(*
SPDX-FileCopyrightText: © 2026 Oleksandr Tiutyk <trofimich@gmail.com>
SPDX-License-Identifier: MIT
License: https://opensource.org/license/mit
*)

(*!
<summary>Represents a named event occurrence without additional payload.</summary>
<description>
Copies its initialization name into instance storage and exposes it through the read-only INamed contract. The
caller must supply a nonempty name. Global uniqueness is not required; each recipient defines how it
recognizes events. Equal names alone do not establish event instance identity. The Event lifetime contract
applies: one instance per occurrence, synchronous borrowed delivery, no retention by recipients and no reset
for reuse as another occurrence. Heap allocation is not required.
</description>
*)

{attribute 'no_explicit_call' := 'do not call this function block directly'}
FUNCTION_BLOCK SimpleEvent EXTENDS Event IMPLEMENTS INamed
VAR_STAT
	//! <summary>Class name shared by all instances of this function block.</summary>
	{attribute 'hide'} 
	_ClassName : STRING := __POUNAME();
END_VAR
VAR
	{attribute 'hide'} 
	_Name : WSTRING;
END_VAR

{attribute 'monitoring' := 'call'}
PROPERTY ClassName : REFERENCE TO STRING
GET
ClassName REF= _ClassName;
END_GET
END_PROPERTY

(*!
<summary>Initializes the event's name; Event initialization associates the optional source.</summary>
<description>
Copies the name into instance storage. The source is borrowed without ownership transfer; the caller must keep
a non-null source alive for the entire event lifetime. The caller must supply a nonempty name; this
precondition is not checked at runtime. Pass both additional initialization arguments explicitly; zero is
allowed for sourceObject.
</description>
*)

//!<param name="sourceObject">Source of the event, or 0 for an event without a specific source.</param>
//!<param name="name">Nonempty name copied into this event instance; global uniqueness is not required.</param>
METHOD FB_init : BOOL
VAR_INPUT
	bInitRetains : BOOL; // TRUE: the retain variables are initialized (reset warm / reset cold)
	bInCopyCode : BOOL;  // TRUE: the instance will be copied to the copy code afterward (online change)
	sourceObject : IObject;
	name : WSTRING;
END_VAR
_Name := name;
END_METHOD

(*!
<summary>Returns a borrowed, read-only view of the event's nonempty name.</summary>
<description>
Requires initialization with a nonempty name. The reference remains usable only while this instance is alive;
callers must not write through it. Recognition rules belong to the recipient, and names need not be globally
unique.
</description>
*)

{attribute 'monitoring' := 'call'}
PROPERTY FINAL Name : REFERENCE TO WSTRING
GET
Name REF= _Name;
END_GET
END_PROPERTY

(*!
<summary>Provides the library namespace used in diagnostics.</summary>
<description>
Borrowed read-only reference to the compiler-initialized library namespace; no ownership transfer.
</description>
*)
{attribute 'monitoring' := 'call'}
PROPERTY NamespaceName : REFERENCE TO STRING
GET
NamespaceName REF= CurrentNamespace.Name;
END_GET
END_PROPERTY

(*!
<summary>Reports the byte size of this concrete instance.</summary>
<description>
Uses XSIZEOF on the instance. Does not include separately allocated payloads or prove that an arbitrary
address is valid.
</description>
*)
{attribute 'monitoring' := 'call'}
PROPERTY SelfSize : ULINT
GET
SelfSize := XSIZEOF(THIS^);
END_GET
END_PROPERTY

END_FUNCTION_BLOCK

(* stored: Version 1.1.0.1
   POU SimpleEvent: Id {6068111a-5f7a-4513-bc9f-2ae69d62cec9}, SpecialFunc None
   Property ClassName: Id {74c80bc7-04ea-415b-b755-fddcf5a7aecd}
   Get Get: Id {0b51e612-0055-4cf8-b992-12a817738a31}
   Method FB_init: Id {95fe79f8-57ab-4f8f-8458-df22c083e6ed}
   Property Name: Id {4cc1da98-6df4-40c6-a0ac-2b058bef2a45}
   Get Get: Id {ad2c60a7-000d-4095-a6d7-745948b89b90}
   Property NamespaceName: Id {1b34e43a-b41f-4a0e-a898-2b2522bb7be9}
   Get Get: Id {3f60aa11-e0bd-4b9d-855a-97e19aaee39b}
   Property SelfSize: Id {f60f572d-0842-4bee-822f-fb69e5ace254}
   Get Get: Id {45257b9e-307e-4ab0-ac78-b362d5465874} *)
